Fanuc KAREL source: KA00044.KL

PROGRAM KA00044
%NOLOCKGROUP
VAR
  SRC: STRING[80]
  DST: JOINTPOS
BEGIN
  SRC = 'A'
  DST = SRC
END KA00044
